{attribute 'Tc2GvlVarNames'}
VAR_GLOBAL
	sgAmsNetId					:STRING := '';						(* AmsNetID of the controller, '' = local netid *)
	lrgActCycleTime				:LREAL;								(* Actual cycle time *)
	// stgSystemTaskInfoArr       		AT%MB32832 :ARRAY[1..4] OF SYSTEMTASKINFOTYPE;
	
	_PlcAppSystemInfo			:PlcAppSystemInfo;
	_PlcTaskSystemInfo			:PlcTaskSystemInfo;	
END_VAR

(* stored: Version 1.1.0.1, ProductVersion 3.1.4024.15
   GVL GVL: Id {fad94044-f1a1-41f5-b5ec-f53828401910} *)
